(* IEC 61131-3 sources: codesys-framework/txt/application/WeVe General (library)/CsvFileLogger/FB_CsvFileLogger, 3 files *)

(* ---- FB_Init.method.st ---- *)
//FB_Init is always available implicitly and it is used primarily for initialization.
//The return value is not evaluated. For a specific influence, you can also declare the
//methods explicitly and provide additional code there with the standard initialization
//code. You can evaluate the return value.
METHOD FB_Init: BOOL
VAR_INPUT
    bInitRetains: BOOL; // TRUE: the retain variables are initialized (reset warm / reset cold)
    bInCopyCode: BOOL;  // TRUE: the instance will be copied to the copy code afterward (online change)

	sFileName 		: STRING(255);			// bv. 'eventlog.csv', relatief tov de bestandsmap van de PLC
	fbTimeStamp 	: I_TimeStampService;	// mag 0 zijn: dan blijft de tijdstempel leeg
END_VAR

// --- BEGIN IMPLEMENTATION ---

// Enkel referenties en waarden bewaren, geen methodes aanroepen
_sFileName 		:= sFileName;
_fbTimeStamp 	:= fbTimeStamp;

(* ---- LogEvent.method.st ---- *)
// Een event loggen. Een tekstlogger gebruikt enkel de tekst (en het level voor de kolom Level);
// ID, bron en payload zitten al in sMessage.
// TRUE = opgenomen in de buffer, FALSE = buffer vol.
METHOD LogEvent : BOOL
VAR_INPUT
	scEvent 		: SC_Event;
	scPayload 		: SC_EventPayload;
	sMessage 		: STRING(GVL_Logger.cMaxMessageLength);
END_VAR

// --- BEGIN IMPLEMENTATION ---

LogEvent := AddEntry(eLevel := scEvent.eEventLevel, sMessage := sMessage);

(* ---- LogMessage.method.st ---- *)
// Vrije tekst loggen, bv. om te debuggen.
// TRUE = opgenomen in de buffer, FALSE = buffer vol.
METHOD LogMessage : BOOL
VAR_INPUT
	eLevel 			: E_EventLevels;
	sMessage 		: STRING(GVL_Logger.cMaxMessageLength);
END_VAR

// --- BEGIN IMPLEMENTATION ---

LogMessage := AddEntry(eLevel := eLevel, sMessage := sMessage);
